(* IEC 61131-3 sources: garage-sweeper/PLC/src/Platform, 3 files *)

(* ---- I_DifferentialDrive.st ---- *)
INTERFACE I_DifferentialDrive
METHOD Execute
METHOD Enable
METHOD Disable
METHOD SetTwist
VAR_INPUT
	desiredTwist : Twist;
END_VAR
PROPERTY LeftWheelPositionInM : LREAL
GET
PROPERTY RightWheelPositionInM : LREAL
GET
PROPERTY IsReady : BOOL
GET

(* ---- DiffDrive.st ---- *)
{attribute 'linkalways'}
{attribute 'no_explicit_call' := 'Use the methods of this class'}
{attribute 'enable_dynamic_creation'}
FUNCTION_BLOCK DiffDrive IMPLEMENTS I_DifferentialDrive
VAR
	leftAxis : I_DriveAxis;
	rightAxis : I_DriveAxis;
	kinematics : DiffDriveKinematics;
END_VAR
METHOD Connect
VAR_INPUT
	left : I_DriveAxis;
	right : I_DriveAxis;
END_VAR
// @impl
leftAxis := left;
rightAxis := right;
END_METHOD
METHOD Execute
// @impl
IF leftAxis = 0 OR rightAxis = 0 THEN
	RETURN;
END_IF
leftAxis.Execute();
rightAxis.Execute();
END_METHOD
METHOD Enable
// @impl
IF leftAxis = 0 OR rightAxis = 0 THEN
	RETURN;
END_IF
leftAxis.Enable();
rightAxis.Enable();
END_METHOD
METHOD Disable
// @impl
IF leftAxis = 0 OR rightAxis = 0 THEN
	RETURN;
END_IF
leftAxis.Disable();
rightAxis.Disable();
END_METHOD
METHOD SetTwist
VAR_INPUT
	desiredTwist : Twist;
END_VAR
VAR
	speeds : WheelSpeeds;
END_VAR
// @impl
IF leftAxis = 0 OR rightAxis = 0 THEN
	RETURN;
END_IF
speeds := kinematics.ToWheelSpeeds(desiredTwist);
leftAxis.SetVelocity(speeds.leftInMPerS);
rightAxis.SetVelocity(speeds.rightInMPerS);
END_METHOD
PROPERTY LeftWheelPositionInM : LREAL
GET
IF leftAxis <> 0 THEN
	LeftWheelPositionInM := leftAxis.PositionInM;
END_IF
END_GET
END_PROPERTY
PROPERTY RightWheelPositionInM : LREAL
GET
IF rightAxis <> 0 THEN
	RightWheelPositionInM := rightAxis.PositionInM;
END_IF
END_GET
END_PROPERTY
PROPERTY IsReady : BOOL
GET
IsReady := leftAxis <> 0 AND_THEN rightAxis <> 0 AND_THEN leftAxis.IsReady AND_THEN rightAxis.IsReady;
END_GET
END_PROPERTY

(* ---- DiffDriveKinematics.st ---- *)
{attribute 'linkalways'}
{attribute 'no_explicit_call' := 'Use the methods of this class'}
{attribute 'enable_dynamic_creation'}
FUNCTION_BLOCK DiffDriveKinematics
METHOD ToWheelSpeeds : WheelSpeeds
VAR_INPUT
	desiredTwist : Twist;
END_VAR
VAR
	speeds : WheelSpeeds;
END_VAR
// @impl
// OPPGAVE M1 (Stian): Gjør robotens fart (twist) om til fart for hvert hjul, i m/s langs hjulbanen.
// Bruk Parameters.trackWidthInM. Hjulradien trengs ikke, den ligger i NC-skaleringen.
// Tips: hvert hjul ligger trackWidth / 2 fra midten. Når roboten roterer med yawRate,
// får hjulet på utsiden ekstra fart lik yawRate * trackWidth / 2.
speeds.leftInMPerS := 0;
speeds.rightInMPerS := 0;
ToWheelSpeeds := speeds;
END_METHOD
METHOD ToBodyMotion : BodyMotion
VAR_INPUT
	leftDeltaInM : LREAL;
	rightDeltaInM : LREAL;
END_VAR
VAR
	motion : BodyMotion;
END_VAR
// @impl
// OPPGAVE M1 (Stian): Gjør hjulenes strekning siden forrige syklus om til robotens strekning og kursendring.
// Den motsatte veien av ToWheelSpeeds: snittet av hjulene gir strekning,
// forskjellen delt på sporvidden gir kursendring.
motion.distanceInM := 0;
motion.headingChangeInRad := 0;
ToBodyMotion := motion;
END_METHOD
